Staubli VAL3: onStart.pgx

program onStart()
  local num l_nResult
  local string l_sKey
  local num l_i
  local num l_nSize
begin

  sUsingLib=toString("",saveData:nLibIndex)
  // l_nResult=trajTemp:libLoad("Disk://data/CustomerLib/lib0/saveTRAJ")
  //  call trajectory:loadTRAJ(0,l_nResult)
  //  if l_nResult!=0
  //    popUpMsg("库加载错误："+toString("",l_nResult))
  //  endIf



  call refreshlist()
  //refresh list
  //  l_sKey=first(trajTemp:tTrajItem)
  //  while l_sKey!=""
  //    sList[size(sList)-1]=l_sKey
  //    insert(sList[size(sList)])
  //    l_sKey=next(trajTemp:tTrajItem[l_sKey])
  //  endWhile

  nPageIndex=0

  if l_nSize>0
    sSelTraj=sList[l_nSize-1]
  else
    sSelTraj=""
  endIf
  //
end
